Fanuc KAREL source: kt00534.KL

-- PROVISIONAL review KL for V770-1; original PC SHA256 9dc475725ed8fce0771b5ccef050d1210cc678b7941207bbcefedb625286aeb5
-- Incomplete behavior may be omitted. Consult companion uncertainty JSON. Do not deploy.
PROGRAM KT00534
%NOLOCKGROUP
-- UNRESOLVED_DECL P1 type=000199
-- UNRESOLVED_DECL P2 type=000101
-- UNRESOLVED_DECL OUT type=000101
BEGIN
  -- UNRESOLVED_PC offsets 5-34; opcodes 49,7E,49,60,4A
  -- UNRESOLVED_PC offsets 39-43; opcodes 7F
END KT00534
